FUNCTION_BLOCK Sensor (* Composite Function Block Type *)
  (* Standard: 61499-2 *)
  (* Version 0.0, 5/26/2016, Andrei, nxtControl GmbH, template *)
  PACKAGE Main;
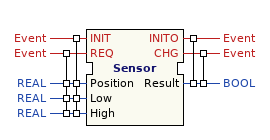
  EVENT_INPUT
    INIT WITH Position, Low, High;
    REQ WITH Position, Low, High; (* Normal Execution Request *)
  END_EVENT
  EVENT_OUTPUT
    INITO WITH Result;
    CHG WITH Result; (* Initialization Confirm *)
  END_EVENT
  VAR_INPUT
    Position : REAL; (* Input event qualifier *)
    Low : REAL;
    High : REAL;
  END_VAR
  VAR_OUTPUT
    Result : BOOL; (* Output event qualifier *)
  END_VAR
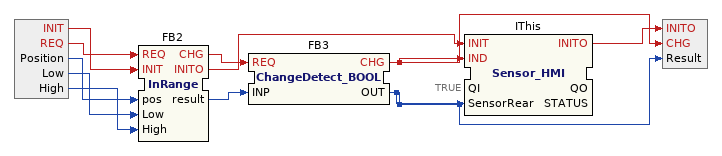
  FBS
    FB2 : InRange;
    IThis : Sensor_HMI(QI := TRUE);
    FB3 : ChangeDetect_BOOL;
  END_FBS
  EVENT_CONNECTIONS
    REQ TO FB2.REQ;
    INIT TO FB2.INIT;
    FB2.CHG TO FB3.REQ;
    FB2.INITO TO IThis.INIT;
    FB3.CHG TO IThis.IND;
    IThis.INITO TO INITO;
    FB3.CHG TO CHG;
  END_CONNECTIONS
  DATA_CONNECTIONS
    Position TO FB2.pos;
    Low TO FB2.Low;
    FB3.OUT TO IThis.SensorRear;
    FB2.result TO FB3.INP;
    FB3.OUT TO Result;
    High TO FB2.High;
  END_CONNECTIONS
END_FUNCTION_BLOCK
